(*
SPDX-FileCopyrightText: © 2026 Oleksandr Tiutyk <trofimich@gmail.com>
SPDX-License-Identifier: MIT
License: https://opensource.org/license/mit
*)

(*!
<summary>Creates generic value descriptors by borrowing, adopting or cloning data.</summary>
<description>
Object cloning requires ICloneable; other cloned values are copied as bytes. Owning modes require permission
to release the stored allocation. Exception objects and their engine-managed clones are unsupported in
user-managed generic collections.
</description>
*)

{attribute 'no_explicit_call' := 'do not call this function block directly'}
PROGRAM GenericValueFactory
VAR_OUTPUT
	GenericValueClassName : STRING := 'GENERIC_VALUE';
END_VAR
VAR
	{attribute 'hide'} 
	_ClassName : STRING := __POUNAME();
END_VAR

{attribute 'monitoring' := 'call'}
PROPERTY ClassName : REFERENCE TO STRING
GET
ClassName REF= _ClassName;
END_GET
END_PROPERTY

(*!
<summary>Creates a generic descriptor from runtime type metadata and the requested memory policy.</summary>
<description>
TYPE_ENUM and TYPE_SUBRANGE are interpreted as unsigned integers of the same byte size; their signedness and
original type identity are not retained. Convert explicitly to a signed integer first when signed numeric
meaning is required. Borrowing a converted variable references that variable, not the original enum/subrange.
The selected memory policy and cloning requirements follow FromParts; borrowed storage must remain alive while
used.
</description>
*)
METHOD FromAny : GENERIC_VALUE
VAR_INPUT
	value : ANY;
	isObject : BOOL;
	memoryManagementBehavior : GENERIC_MEMORY_MANAGEMENT_BEHAVIOR;
END_VAR
FromAny := FromAnyType(
	value := value,
	isObject := isObject,
	memoryManagementBehavior := memoryManagementBehavior
);
END_METHOD

(*!
<summary>Creates a generic descriptor from runtime type metadata and the requested memory policy.</summary>
<description>
TYPE_ENUM and TYPE_SUBRANGE are interpreted as unsigned integers of the same byte size; their signedness and
original type identity are not retained. Convert explicitly to a signed integer first when signed numeric
meaning is required. Borrowing a converted variable references that variable, not the original enum/subrange.
The selected memory policy and cloning requirements follow FromParts; borrowed storage must remain alive while
used.
</description>
*)
METHOD FromAnyType : GENERIC_VALUE
VAR_INPUT
	value : __SYSTEM.AnyType;
	isObject : BOOL;
	memoryManagementBehavior : GENERIC_MEMORY_MANAGEMENT_BEHAVIOR;
END_VAR
FromAnyType := FromParts(
        	genericTypeClass := GenericTypeClassConvertor.GetGenericTypeClassBySystemAnyType(systemAnyType := value, isObject := isObject),
        	address := value.pValue,
        	size := TO_ULINT(value.diSize),
        	memoryManagementBehavior := memoryManagementBehavior
        );
END_METHOD

(*!
<summary>Borrows existing storage as a BOOLEAN descriptor.</summary>
<description>
Does not copy or own the payload. The caller keeps the source alive and its representation stable while the
descriptor is used. Size is the byte size of the source variable.
</description>
*)
METHOD FromBoolReference : GENERIC_VALUE
VAR_IN_OUT
	value : BOOL;
END_VAR
FromBoolReference := FromParts(
        	genericTypeClass := GENERIC_TYPE_CLASS.BOOLEAN,
        	address := ADR(value),
        	size := XSIZEOF(value),
        	memoryManagementBehavior := GENERIC_MEMORY_MANAGEMENT_BEHAVIOR.STORE_ORIGINAL_REFERENCE_AND_NOT_OWNS_MEMORY
        );
END_METHOD

(*!
<summary>Creates an owned snapshot of a BOOL value.</summary>
<description>
The result is independent of the input storage; release it or transfer ownership exactly once. Allocation
failure uses the framework terminal allocation path. Uses FromAny cloning; the source value is not modified.
</description>
*)
METHOD FromBoolValue : GENERIC_VALUE
VAR_INPUT
	value : BOOL;
END_VAR
FromBoolValue := FromAny(
	value := value,
	isObject := FALSE,
	memoryManagementBehavior := GENERIC_MEMORY_MANAGEMENT_BEHAVIOR.CLONE_ORIGINAL_VALUE_AND_OWNS_MEMORY
);
END_METHOD

(*!
<summary>Borrows existing storage as a UINT_8 descriptor.</summary>
<description>
Does not copy or own the payload. The caller keeps the source alive and its representation stable while the
descriptor is used. Size is the byte size of the source variable.
</description>
*)
METHOD FromByteReference : GENERIC_VALUE
VAR_IN_OUT
	value : BYTE;
END_VAR
FromByteReference := FromParts(
        	genericTypeClass := GENERIC_TYPE_CLASS.UINT_8,
        	address := ADR(value),
        	size := XSIZEOF(value),
        	memoryManagementBehavior := GENERIC_MEMORY_MANAGEMENT_BEHAVIOR.STORE_ORIGINAL_REFERENCE_AND_NOT_OWNS_MEMORY
        );
END_METHOD

(*!
<summary>Creates an owned snapshot of a BYTE value.</summary>
<description>
The result is independent of the input storage; release it or transfer ownership exactly once. Allocation
failure uses the framework terminal allocation path. Uses FromAny cloning; the source value is not modified.
</description>
*)
METHOD FromByteValue : GENERIC_VALUE
VAR_INPUT
	value : BYTE;
END_VAR
FromByteValue := FromAny(
	value := value,
	isObject := FALSE,
	memoryManagementBehavior := GENERIC_MEMORY_MANAGEMENT_BEHAVIOR.CLONE_ORIGINAL_VALUE_AND_OWNS_MEMORY
);
END_METHOD

(*!
<summary>Borrows existing storage as a DATE_AND_TIME_32 descriptor.</summary>
<description>
Does not copy or own the payload. The caller keeps the source alive and its representation stable while the
descriptor is used. Size is the byte size of the source variable.
</description>
*)
METHOD FromDateAndTimeReference : GENERIC_VALUE
VAR_IN_OUT
	value : DATE_AND_TIME;
END_VAR
FromDateAndTimeReference := FromParts(
        	genericTypeClass := GENERIC_TYPE_CLASS.DATE_AND_TIME_32,
        	address := ADR(value),
        	size := XSIZEOF(value),
        	memoryManagementBehavior := GENERIC_MEMORY_MANAGEMENT_BEHAVIOR.STORE_ORIGINAL_REFERENCE_AND_NOT_OWNS_MEMORY
        );
END_METHOD

(*!
<summary>Creates an owned snapshot of a DATE_AND_TIME value.</summary>
<description>
The result is independent of the input storage; release it or transfer ownership exactly once. Allocation
failure uses the framework terminal allocation path. Uses FromAny cloning; the source value is not modified.
</description>
*)
METHOD FromDateAndTimeValue : GENERIC_VALUE
VAR_INPUT
	value : DATE_AND_TIME;
END_VAR
FromDateAndTimeValue := FromAny(
	value := value,
	isObject := FALSE,
	memoryManagementBehavior := GENERIC_MEMORY_MANAGEMENT_BEHAVIOR.CLONE_ORIGINAL_VALUE_AND_OWNS_MEMORY
);
END_METHOD

(*!
<summary>Borrows existing storage as a DATE_32 descriptor.</summary>
<description>
Does not copy or own the payload. The caller keeps the source alive and its representation stable while the
descriptor is used. Size is the byte size of the source variable.
</description>
*)
METHOD FromDateReference : GENERIC_VALUE
VAR_IN_OUT
	value : DATE;
END_VAR
FromDateReference := FromParts(
        	genericTypeClass := GENERIC_TYPE_CLASS.DATE_32,
        	address := ADR(value),
        	size := XSIZEOF(value),
        	memoryManagementBehavior := GENERIC_MEMORY_MANAGEMENT_BEHAVIOR.STORE_ORIGINAL_REFERENCE_AND_NOT_OWNS_MEMORY
        );
END_METHOD

(*!
<summary>Creates an owned snapshot of a DATE value.</summary>
<description>
The result is independent of the input storage; release it or transfer ownership exactly once. Allocation
failure uses the framework terminal allocation path. Uses FromAny cloning; the source value is not modified.
</description>
*)
METHOD FromDateValue : GENERIC_VALUE
VAR_INPUT
	value : DATE;
END_VAR
FromDateValue := FromAny(
	value := value,
	isObject := FALSE,
	memoryManagementBehavior := GENERIC_MEMORY_MANAGEMENT_BEHAVIOR.CLONE_ORIGINAL_VALUE_AND_OWNS_MEMORY
);
END_METHOD

(*!
<summary>Borrows existing storage as a INT_32 descriptor.</summary>
<description>
Does not copy or own the payload. The caller keeps the source alive and its representation stable while the
descriptor is used. Size is the byte size of the source variable.
</description>
*)
METHOD FromDIntReference : GENERIC_VALUE
VAR_IN_OUT
	value : DINT;
END_VAR
FromDIntReference := FromParts(
        	genericTypeClass := GENERIC_TYPE_CLASS.INT_32,
        	address := ADR(value),
        	size := XSIZEOF(value),
        	memoryManagementBehavior := GENERIC_MEMORY_MANAGEMENT_BEHAVIOR.STORE_ORIGINAL_REFERENCE_AND_NOT_OWNS_MEMORY
        );
END_METHOD

(*!
<summary>Creates an owned snapshot of a DINT value.</summary>
<description>
The result is independent of the input storage; release it or transfer ownership exactly once. Allocation
failure uses the framework terminal allocation path. Uses FromAny cloning; the source value is not modified.
</description>
*)
METHOD FromDIntValue : GENERIC_VALUE
VAR_INPUT
	value : DINT;
END_VAR
FromDIntValue := FromAny(
	value := value,
	isObject := FALSE,
	memoryManagementBehavior := GENERIC_MEMORY_MANAGEMENT_BEHAVIOR.CLONE_ORIGINAL_VALUE_AND_OWNS_MEMORY
);
END_METHOD

(*!
<summary>Borrows existing storage as a UINT_32 descriptor.</summary>
<description>
Does not copy or own the payload. The caller keeps the source alive and its representation stable while the
descriptor is used. Size is the byte size of the source variable.
</description>
*)
METHOD FromDWordReference : GENERIC_VALUE
VAR_IN_OUT
	value : DWORD;
END_VAR
FromDWordReference := FromParts(
        	genericTypeClass := GENERIC_TYPE_CLASS.UINT_32,
        	address := ADR(value),
        	size := XSIZEOF(value),
        	memoryManagementBehavior := GENERIC_MEMORY_MANAGEMENT_BEHAVIOR.STORE_ORIGINAL_REFERENCE_AND_NOT_OWNS_MEMORY
        );
END_METHOD

(*!
<summary>Creates an owned snapshot of a DWORD value.</summary>
<description>
The result is independent of the input storage; release it or transfer ownership exactly once. Allocation
failure uses the framework terminal allocation path. Uses FromAny cloning; the source value is not modified.
</description>
*)
METHOD FromDWordValue : GENERIC_VALUE
VAR_INPUT
	value : DWORD;
END_VAR
FromDWordValue := FromAny(
	value := value,
	isObject := FALSE,
	memoryManagementBehavior := GENERIC_MEMORY_MANAGEMENT_BEHAVIOR.CLONE_ORIGINAL_VALUE_AND_OWNS_MEMORY
);
END_METHOD

(*!
<summary>Borrows existing storage as a INT_16 descriptor.</summary>
<description>
Does not copy or own the payload. The caller keeps the source alive and its representation stable while the
descriptor is used. Size is the byte size of the source variable.
</description>
*)
METHOD FromIntReference : GENERIC_VALUE
VAR_IN_OUT
	value : INT;
END_VAR
FromIntReference := FromParts(
        	genericTypeClass := GENERIC_TYPE_CLASS.INT_16,
        	address := ADR(value),
        	size := XSIZEOF(value),
        	memoryManagementBehavior := GENERIC_MEMORY_MANAGEMENT_BEHAVIOR.STORE_ORIGINAL_REFERENCE_AND_NOT_OWNS_MEMORY
        );
END_METHOD

(*!
<summary>Creates an owned snapshot of a INT value.</summary>
<description>
The result is independent of the input storage; release it or transfer ownership exactly once. Allocation
failure uses the framework terminal allocation path. Uses FromAny cloning; the source value is not modified.
</description>
*)
METHOD FromIntValue : GENERIC_VALUE
VAR_INPUT
	value : INT;
END_VAR
FromIntValue := FromAny(
	value := value,
	isObject := FALSE,
	memoryManagementBehavior := GENERIC_MEMORY_MANAGEMENT_BEHAVIOR.CLONE_ORIGINAL_VALUE_AND_OWNS_MEMORY
);
END_METHOD

(*!
<summary>Creates a non-owning descriptor for an existing object.</summary>
<description>
Null input raises ArgumentNotSpecifiedException. Uses the live object SelfAddress and SelfSize; does not clone
or retain ownership. The object must outlive all uses of the result.
</description>
*)
METHOD FromIObjectReference : GENERIC_VALUE
VAR_INPUT
	instance : IObject;
END_VAR
IF instance = 0 THEN
	Exceptions.ThrowArgumentNotSpecified(
		sourceNamespaceName := NamespaceName,
		sourceClassName := ClassName,
		sourcePOUName := __POUNAME(),
		sourcePosition := __POSITION(),
		argumentName := 'instance'
	);
END_IF

FromIObjectReference := FromParts(
		genericTypeClass := GENERIC_TYPE_CLASS.OBJECT,
		address := instance.SelfAddress,
		size := instance.SelfSize,
		memoryManagementBehavior := GENERIC_MEMORY_MANAGEMENT_BEHAVIOR.STORE_ORIGINAL_REFERENCE_AND_NOT_OWNS_MEMORY
	);
END_METHOD

(*!
<summary>Creates an owning descriptor for a clone of an object.</summary>
<description>
Null input raises ArgumentNotSpecifiedException. Uses the FromParts object-clone contract: a suitable
independent ICloneable result is required; failure raises an exception. The caller must release or transfer
the result exactly once. Task-managed exception clones are not supported as owned generic values.
</description>
*)
METHOD FromIObjectValue : GENERIC_VALUE 
VAR_INPUT
	instance : IObject;
END_VAR
IF instance = 0 THEN
	Exceptions.ThrowArgumentNotSpecified(
		sourceNamespaceName := NamespaceName,
		sourceClassName := ClassName,
		sourcePOUName := __POUNAME(),
		sourcePosition := __POSITION(),
		argumentName := 'instance'
	);
END_IF

FromIObjectValue := FromParts(
		genericTypeClass := GENERIC_TYPE_CLASS.OBJECT,
		address := instance.SelfAddress,
		size := instance.SelfSize,
		memoryManagementBehavior := GENERIC_MEMORY_MANAGEMENT_BEHAVIOR.CLONE_ORIGINAL_VALUE_AND_OWNS_MEMORY
	);
END_METHOD

(*!
<summary>Creates a borrowed generic descriptor for an LDATE_AND_TIME variable.</summary>
<description>
Preserves the DATE_AND_TIME_64 category and references the original variable without copying or allocating
storage. The caller keeps the variable alive while the descriptor is used; ownership is not transferred.
</description>
*)
//!<param name="value">Variable whose storage is borrowed by the returned descriptor.</param>
METHOD FromLDateAndTimeReference : GENERIC_VALUE
VAR_IN_OUT
	value : LDATE_AND_TIME;
END_VAR
FromLDateAndTimeReference := FromParts(
        	genericTypeClass := GENERIC_TYPE_CLASS.DATE_AND_TIME_64,
        	address := ADR(value),
        	size := XSIZEOF(value),
        	memoryManagementBehavior := GENERIC_MEMORY_MANAGEMENT_BEHAVIOR.STORE_ORIGINAL_REFERENCE_AND_NOT_OWNS_MEMORY
        );
END_METHOD

(*!
<summary>Creates an owned snapshot of a LDATE_AND_TIME value.</summary>
<description>
The result is independent of the input storage; release it or transfer ownership exactly once. Allocation
failure uses the framework terminal allocation path. Uses FromAny cloning; the source value is not modified.
</description>
*)
METHOD FromLDateAndTimeValue : GENERIC_VALUE
VAR_INPUT
	value : LDATE_AND_TIME;
END_VAR
FromLDateAndTimeValue := FromAny(
	value := value,
	isObject := FALSE,
	memoryManagementBehavior := GENERIC_MEMORY_MANAGEMENT_BEHAVIOR.CLONE_ORIGINAL_VALUE_AND_OWNS_MEMORY
);
END_METHOD

(*!
<summary>Creates a borrowed generic descriptor for an LDATE variable.</summary>
<description>
Preserves the DATE_64 category and references the original variable without copying or allocating storage. The
caller keeps the variable alive while the descriptor is used; ownership is not transferred.
</description>
*)
//!<param name="value">Variable whose storage is borrowed by the returned descriptor.</param>
METHOD FromLDateReference : GENERIC_VALUE
VAR_IN_OUT
	value : LDATE;
END_VAR
FromLDateReference := FromParts(
        	genericTypeClass := GENERIC_TYPE_CLASS.DATE_64,
        	address := ADR(value),
        	size := XSIZEOF(value),
        	memoryManagementBehavior := GENERIC_MEMORY_MANAGEMENT_BEHAVIOR.STORE_ORIGINAL_REFERENCE_AND_NOT_OWNS_MEMORY
        );
END_METHOD

(*!
<summary>Creates an owned snapshot of a LDATE value.</summary>
<description>
The result is independent of the input storage; release it or transfer ownership exactly once. Allocation
failure uses the framework terminal allocation path. Uses FromAny cloning; the source value is not modified.
</description>
*)
METHOD FromLDateValue : GENERIC_VALUE
VAR_INPUT
	value : LDATE;
END_VAR
FromLDateValue := FromAny(
	value := value,
	isObject := FALSE,
	memoryManagementBehavior := GENERIC_MEMORY_MANAGEMENT_BEHAVIOR.CLONE_ORIGINAL_VALUE_AND_OWNS_MEMORY
);
END_METHOD

(*!
<summary>Borrows existing storage as a INT_64 descriptor.</summary>
<description>
Does not copy or own the payload. The caller keeps the source alive and its representation stable while the
descriptor is used. Size is the byte size of the source variable.
</description>
*)
METHOD FromLIntReference : GENERIC_VALUE
VAR_IN_OUT
	value : LINT;
END_VAR
FromLIntReference := FromParts(
        	genericTypeClass := GENERIC_TYPE_CLASS.INT_64,
        	address := ADR(value),
        	size := XSIZEOF(value),
        	memoryManagementBehavior := GENERIC_MEMORY_MANAGEMENT_BEHAVIOR.STORE_ORIGINAL_REFERENCE_AND_NOT_OWNS_MEMORY
        );
END_METHOD

(*!
<summary>Creates an owned snapshot of a LINT value.</summary>
<description>
The result is independent of the input storage; release it or transfer ownership exactly once. Allocation
failure uses the framework terminal allocation path. Uses FromAny cloning; the source value is not modified.
</description>
*)
METHOD FromLIntValue : GENERIC_VALUE
VAR_INPUT
	value : LINT;
END_VAR
FromLIntValue := FromAny(
	value := value,
	isObject := FALSE,
	memoryManagementBehavior := GENERIC_MEMORY_MANAGEMENT_BEHAVIOR.CLONE_ORIGINAL_VALUE_AND_OWNS_MEMORY
);
END_METHOD

(*!
<summary>Borrows existing storage as a REAL_64 descriptor.</summary>
<description>
Does not copy or own the payload. The caller keeps the source alive and its representation stable while the
descriptor is used. Size is the byte size of the source variable.
</description>
*)
METHOD FromLRealReference : GENERIC_VALUE
VAR_IN_OUT
	value : LREAL;
END_VAR
FromLRealReference := FromParts(
        	genericTypeClass := GENERIC_TYPE_CLASS.REAL_64,
        	address := ADR(value),
        	size := XSIZEOF(value),
        	memoryManagementBehavior := GENERIC_MEMORY_MANAGEMENT_BEHAVIOR.STORE_ORIGINAL_REFERENCE_AND_NOT_OWNS_MEMORY
        );
END_METHOD

(*!
<summary>Creates an owned snapshot of a LREAL value.</summary>
<description>
The result is independent of the input storage; release it or transfer ownership exactly once. Allocation
failure uses the framework terminal allocation path. Uses FromAny cloning; the source value is not modified.
</description>
*)
METHOD FromLRealValue : GENERIC_VALUE
VAR_INPUT
	value : LREAL;
END_VAR
FromLRealValue := FromAny(
	value := value,
	isObject := FALSE,
	memoryManagementBehavior := GENERIC_MEMORY_MANAGEMENT_BEHAVIOR.CLONE_ORIGINAL_VALUE_AND_OWNS_MEMORY
);
END_METHOD

(*!
<summary>Creates a borrowed generic descriptor for an LTIME_OF_DAY variable.</summary>
<description>
Preserves the TIME_OF_DAY_64 category and references the original variable without copying or allocating
storage. The caller keeps the variable alive while the descriptor is used; ownership is not transferred.
</description>
*)
//!<param name="value">Variable whose storage is borrowed by the returned descriptor.</param>
METHOD FromLTimeOfDayReference : GENERIC_VALUE
VAR_IN_OUT
	value : LTIME_OF_DAY;
END_VAR
FromLTimeOfDayReference := FromParts(
        	genericTypeClass := GENERIC_TYPE_CLASS.TIME_OF_DAY_64,
        	address := ADR(value),
        	size := XSIZEOF(value),
        	memoryManagementBehavior := GENERIC_MEMORY_MANAGEMENT_BEHAVIOR.STORE_ORIGINAL_REFERENCE_AND_NOT_OWNS_MEMORY
        );
END_METHOD

(*!
<summary>Creates an owned snapshot of a LTIME_OF_DAY value.</summary>
<description>
The result is independent of the input storage; release it or transfer ownership exactly once. Allocation
failure uses the framework terminal allocation path. Uses FromAny cloning; the source value is not modified.
</description>
*)
METHOD FromLTimeOfDayValue : GENERIC_VALUE
VAR_INPUT
	value : LTIME_OF_DAY;
END_VAR
FromLTimeOfDayValue := FromAny(
	value := value,
	isObject := FALSE,
	memoryManagementBehavior := GENERIC_MEMORY_MANAGEMENT_BEHAVIOR.CLONE_ORIGINAL_VALUE_AND_OWNS_MEMORY
);
END_METHOD

(*!
<summary>Creates a borrowed generic descriptor for an LTIME variable.</summary>
<description>
Preserves the TIME_64 category and references the original variable without copying or allocating storage. The
caller keeps the variable alive while the descriptor is used; ownership is not transferred.
</description>
*)
//!<param name="value">Variable whose storage is borrowed by the returned descriptor.</param>
METHOD FromLTimeReference : GENERIC_VALUE
VAR_IN_OUT
	value : LTIME;
END_VAR
FromLTimeReference := FromParts(
        	genericTypeClass := GENERIC_TYPE_CLASS.TIME_64,
        	address := ADR(value),
        	size := XSIZEOF(value),
        	memoryManagementBehavior := GENERIC_MEMORY_MANAGEMENT_BEHAVIOR.STORE_ORIGINAL_REFERENCE_AND_NOT_OWNS_MEMORY
        );
END_METHOD

(*!
<summary>Creates an owned snapshot of a LTIME value.</summary>
<description>
The result is independent of the input storage; release it or transfer ownership exactly once. Allocation
failure uses the framework terminal allocation path. Uses FromAny cloning; the source value is not modified.
</description>
*)
METHOD FromLTimeValue : GENERIC_VALUE
VAR_INPUT
	value : LTIME;
END_VAR
FromLTimeValue := FromAny(
	value := value,
	isObject := FALSE,
	memoryManagementBehavior := GENERIC_MEMORY_MANAGEMENT_BEHAVIOR.CLONE_ORIGINAL_VALUE_AND_OWNS_MEMORY
);
END_METHOD

(*!
<summary>Borrows existing storage as a UINT_64 descriptor.</summary>
<description>
Does not copy or own the payload. The caller keeps the source alive and its representation stable while the
descriptor is used. Size is the byte size of the source variable.
</description>
*)
METHOD FromLWordReference : GENERIC_VALUE
VAR_IN_OUT
	value : LWORD;
END_VAR
FromLWordReference := FromParts(
        	genericTypeClass := GENERIC_TYPE_CLASS.UINT_64,
        	address := ADR(value),
        	size := XSIZEOF(value),
        	memoryManagementBehavior := GENERIC_MEMORY_MANAGEMENT_BEHAVIOR.STORE_ORIGINAL_REFERENCE_AND_NOT_OWNS_MEMORY
        );
END_METHOD

(*!
<summary>Creates an owned snapshot of a LWORD value.</summary>
<description>
The result is independent of the input storage; release it or transfer ownership exactly once. Allocation
failure uses the framework terminal allocation path. Uses FromAny cloning; the source value is not modified.
</description>
*)
METHOD FromLWordValue : GENERIC_VALUE
VAR_INPUT
	value : LWORD;
END_VAR
FromLWordValue := FromAny(
	value := value,
	isObject := FALSE,
	memoryManagementBehavior := GENERIC_MEMORY_MANAGEMENT_BEHAVIOR.CLONE_ORIGINAL_VALUE_AND_OWNS_MEMORY
);
END_METHOD

(*!
<summary>Creates a non-owning descriptor for an existing object.</summary>
<description>
Null input raises ArgumentNotSpecifiedException. Uses the live object SelfAddress and SelfSize; does not clone
or retain ownership. The object must outlive all uses of the result.
</description>
*)
METHOD FromObjectReference : GENERIC_VALUE
VAR_INPUT
	instance : REFERENCE TO Object;
END_VAR
IF NOT __ISVALIDREF(instance) THEN
	Exceptions.ThrowArgumentNotSpecified(
		sourceNamespaceName := NamespaceName,
		sourceClassName := ClassName,
		sourcePOUName := __POUNAME(),
		sourcePosition := __POSITION(),
		argumentName := 'instance'
	);
END_IF

FromObjectReference := FromParts(
		genericTypeClass := GENERIC_TYPE_CLASS.OBJECT,
		address := instance.SelfAddress,
		size := instance.SelfSize,
		memoryManagementBehavior := GENERIC_MEMORY_MANAGEMENT_BEHAVIOR.STORE_ORIGINAL_REFERENCE_AND_NOT_OWNS_MEMORY
	);
END_METHOD

(*!
<summary>Creates an owning generic descriptor for a clone of the supplied object.</summary>
<description>
Requires a live object implementing ICloneable whose clone may be released by the owner of the returned
descriptor. Throws ArgumentNotSpecifiedException for a null reference or NotSupportedException when ICloneable
is absent. The original object is not adopted.
</description>
*)
//!<param name="instance">Object to clone through ICloneable.</param>
METHOD FromObjectValue : GENERIC_VALUE 
VAR_INPUT
	instance : REFERENCE TO Object;
END_VAR
IF NOT __ISVALIDREF(instance) THEN
	Exceptions.ThrowArgumentNotSpecified(
		sourceNamespaceName := NamespaceName,
		sourceClassName := ClassName,
		sourcePOUName := __POUNAME(),
		sourcePosition := __POSITION(),
		argumentName := 'instance'
	);
END_IF

FromObjectValue := FromParts(
		genericTypeClass := GENERIC_TYPE_CLASS.OBJECT,
		address := instance.SelfAddress,
		size := instance.SelfSize,
		memoryManagementBehavior := GENERIC_MEMORY_MANAGEMENT_BEHAVIOR.CLONE_ORIGINAL_VALUE_AND_OWNS_MEMORY
	);
END_METHOD

(*!
<summary>Creates a generic value from a type, address, size and memory-management policy.</summary>
<description>
Owning modes require permission to release the stored allocation, including any result returned by Clone. In
clone mode, OBJECT requires ICloneable; otherwise NotSupportedException is raised. Clone must return a
non-null object on success and raise an exception on failure; its exceptions propagate. Failure to allocate a
byte copy invokes the terminal DynamicMemoryManager.RaiseAllocationFailure mechanism. Other type categories
are copied as bytes, without recursively cloning referenced resources. For a nonempty byte copy, size above
UnsignedInt32.MAX_VALUE raises ArgumentOutOfRangeException before allocation or conversion to UDINT. Exception
objects and their engine-managed clones are not supported by user-managed generic collections. Their lifetime
ends at cycle cleanup; use ERROR to retain an error as state.
</description>
*)
METHOD FromParts : GENERIC_VALUE
VAR_INPUT
	genericTypeClass : GENERIC_TYPE_CLASS;
	address : POINTER TO BYTE;
	size : ULINT;
	memoryManagementBehavior : GENERIC_MEMORY_MANAGEMENT_BEHAVIOR;
END_VAR
VAR
	newAddress : POINTER TO BYTE;

	objectPointer : POINTER TO Object;
	cloneable : ICloneable;
	clone : IObject;

END_VAR
IF address = 0 OR_ELSE size <= 0 THEN
	RETURN;
END_IF

CASE memoryManagementBehavior OF
	GENERIC_MEMORY_MANAGEMENT_BEHAVIOR.CLONE_ORIGINAL_VALUE_AND_OWNS_MEMORY:
		IF genericTypeClass = GENERIC_TYPE_CLASS.OBJECT THEN
			objectPointer := address;

			IF NOT __QUERYINTERFACE(objectPointer^, cloneable) THEN
				Exceptions.ThrowNotSupported(
					sourceNamespaceName := NamespaceName,
					sourceClassName := ClassName,
					sourcePOUName := __POUNAME(),
					sourcePosition := __POSITION(),
					message := "Object cloning requires ICloneable."
				);
			END_IF

			clone := cloneable.Clone();
			newAddress := clone.SelfAddress;	
		ELSE
			IF size > TO_ULINT(UnsignedInt32.MAX_VALUE) THEN
				Exceptions.ThrowArgumentOutOfRange(
					sourceNamespaceName := NamespaceName,
					sourceClassName := ClassName,
					sourcePOUName := __POUNAME(),
					sourcePosition := __POSITION(),
					argumentName := 'size',
					argumentValue := size
				);
			END_IF

			newAddress := __NEW(BYTE, TO_UDINT(size));

			IF newAddress = 0 THEN
				DynamicMemoryManager.RaiseAllocationFailure();
			END_IF

			Tc2_System.MEMCPY(destAddr := newAddress, srcAddr := address, n := TO_UDINT(size));
		END_IF

		FromParts.Assign(genericTypeClass := genericTypeClass, address := newAddress, size := size, isMemoryOwner := TRUE);
	
	GENERIC_MEMORY_MANAGEMENT_BEHAVIOR.STORE_ORIGINAL_REFERENCE_AND_NOT_OWNS_MEMORY:
		FromParts.Assign(genericTypeClass := genericTypeClass, address := address, size := size, isMemoryOwner := FALSE);
	
	GENERIC_MEMORY_MANAGEMENT_BEHAVIOR.STORE_ORIGINAL_REFERENCE_AND_OWNS_MEMORY:
		FromParts.Assign(genericTypeClass := genericTypeClass, address := address, size := size, isMemoryOwner := TRUE);
END_CASE
END_METHOD

(*!
<summary>Borrows existing storage as a REAL_32 descriptor.</summary>
<description>
Does not copy or own the payload. The caller keeps the source alive and its representation stable while the
descriptor is used. Size is the byte size of the source variable.
</description>
*)
METHOD FromRealReference : GENERIC_VALUE
VAR_IN_OUT
	value : REAL;
END_VAR
FromRealReference := FromParts(
        	genericTypeClass := GENERIC_TYPE_CLASS.REAL_32,
        	address := ADR(value),
        	size := XSIZEOF(value),
        	memoryManagementBehavior := GENERIC_MEMORY_MANAGEMENT_BEHAVIOR.STORE_ORIGINAL_REFERENCE_AND_NOT_OWNS_MEMORY
        );
END_METHOD

(*!
<summary>Creates an owned snapshot of a REAL value.</summary>
<description>
The result is independent of the input storage; release it or transfer ownership exactly once. Allocation
failure uses the framework terminal allocation path. Uses FromAny cloning; the source value is not modified.
</description>
*)
METHOD FromRealValue : GENERIC_VALUE
VAR_INPUT
	value : REAL;
END_VAR
FromRealValue := FromAny(
	value := value,
	isObject := FALSE,
	memoryManagementBehavior := GENERIC_MEMORY_MANAGEMENT_BEHAVIOR.CLONE_ORIGINAL_VALUE_AND_OWNS_MEMORY
);
END_METHOD

(*!
<summary>Borrows existing storage as a INT_8 descriptor.</summary>
<description>
Does not copy or own the payload. The caller keeps the source alive and its representation stable while the
descriptor is used. Size is the byte size of the source variable.
</description>
*)
METHOD FromSIntReference : GENERIC_VALUE
VAR_IN_OUT
	value : SINT;
END_VAR
FromSIntReference := FromParts(
        	genericTypeClass := GENERIC_TYPE_CLASS.INT_8,
        	address := ADR(value),
        	size := XSIZEOF(value),
        	memoryManagementBehavior := GENERIC_MEMORY_MANAGEMENT_BEHAVIOR.STORE_ORIGINAL_REFERENCE_AND_NOT_OWNS_MEMORY
        );
END_METHOD

(*!
<summary>Creates an owned snapshot of a SINT value.</summary>
<description>
The result is independent of the input storage; release it or transfer ownership exactly once. Allocation
failure uses the framework terminal allocation path. Uses FromAny cloning; the source value is not modified.
</description>
*)
METHOD FromSIntValue : GENERIC_VALUE
VAR_INPUT
	value : SINT;
END_VAR
FromSIntValue := FromAny(
	value := value,
	isObject := FALSE,
	memoryManagementBehavior := GENERIC_MEMORY_MANAGEMENT_BEHAVIOR.CLONE_ORIGINAL_VALUE_AND_OWNS_MEMORY
);
END_METHOD

(*!
<summary>Borrows existing storage as a STRING_8 descriptor.</summary>
<description>
Does not copy or own the payload. The caller keeps the source alive and its representation stable while the
descriptor is used. Size records the current text including its terminator, not the full declared buffer
capacity.
</description>
*)
METHOD FromStringReference : GENERIC_VALUE
VAR_IN_OUT CONSTANT
	value : STRING;
END_VAR
FromStringReference := FromParts(
	genericTypeClass := GENERIC_TYPE_CLASS.STRING_8,
	address := ADR(value),
	size := Strings.GetActualSize(value := value),
	memoryManagementBehavior := GENERIC_MEMORY_MANAGEMENT_BEHAVIOR.STORE_ORIGINAL_REFERENCE_AND_NOT_OWNS_MEMORY
);
END_METHOD

(*!
<summary>Creates an owned snapshot of a STRING value.</summary>
<description>
The result is independent of the input storage; release it or transfer ownership exactly once. Allocation
failure uses the framework terminal allocation path. Copies current text including its terminator, not unused
buffer capacity.
</description>
*)
METHOD FromStringValue : GENERIC_VALUE
VAR_IN_OUT CONSTANT
	value : STRING;
END_VAR
FromStringValue := FromParts(
        	genericTypeClass := GENERIC_TYPE_CLASS.STRING_8,
        	address := ADR(value),
        	size := Strings.GetActualSize(value := value),
        	memoryManagementBehavior := GENERIC_MEMORY_MANAGEMENT_BEHAVIOR.CLONE_ORIGINAL_VALUE_AND_OWNS_MEMORY
        );
END_METHOD

(*!
<summary>Borrows existing storage as a TIME_OF_DAY_32 descriptor.</summary>
<description>
Does not copy or own the payload. The caller keeps the source alive and its representation stable while the
descriptor is used. Size is the byte size of the source variable.
</description>
*)
METHOD FromTimeOfDayReference : GENERIC_VALUE
VAR_IN_OUT
	value : TIME_OF_DAY;
END_VAR
FromTimeOfDayReference := FromParts(
        	genericTypeClass := GENERIC_TYPE_CLASS.TIME_OF_DAY_32,
        	address := ADR(value),
        	size := XSIZEOF(value),
        	memoryManagementBehavior := GENERIC_MEMORY_MANAGEMENT_BEHAVIOR.STORE_ORIGINAL_REFERENCE_AND_NOT_OWNS_MEMORY
        );
END_METHOD

(*!
<summary>Creates an owned snapshot of a TIME_OF_DAY value.</summary>
<description>
The result is independent of the input storage; release it or transfer ownership exactly once. Allocation
failure uses the framework terminal allocation path. Uses FromAny cloning; the source value is not modified.
</description>
*)
METHOD FromTimeOfDayValue : GENERIC_VALUE
VAR_INPUT
	value : TIME_OF_DAY;
END_VAR
FromTimeOfDayValue := FromAny(
	value := value,
	isObject := FALSE,
	memoryManagementBehavior := GENERIC_MEMORY_MANAGEMENT_BEHAVIOR.CLONE_ORIGINAL_VALUE_AND_OWNS_MEMORY
);
END_METHOD

(*!
<summary>Borrows existing storage as a TIME_32 descriptor.</summary>
<description>
Does not copy or own the payload. The caller keeps the source alive and its representation stable while the
descriptor is used. Size is the byte size of the source variable.
</description>
*)
METHOD FromTimeReference : GENERIC_VALUE
VAR_IN_OUT
	value : TIME;
END_VAR
FromTimeReference := FromParts(
        	genericTypeClass := GENERIC_TYPE_CLASS.TIME_32,
        	address := ADR(value),
        	size := XSIZEOF(value),
        	memoryManagementBehavior := GENERIC_MEMORY_MANAGEMENT_BEHAVIOR.STORE_ORIGINAL_REFERENCE_AND_NOT_OWNS_MEMORY
        );
END_METHOD

(*!
<summary>Creates an owned snapshot of a TIME value.</summary>
<description>
The result is independent of the input storage; release it or transfer ownership exactly once. Allocation
failure uses the framework terminal allocation path. Uses FromAny cloning; the source value is not modified.
</description>
*)
METHOD FromTimeValue : GENERIC_VALUE
VAR_INPUT
	value : TIME;
END_VAR
FromTimeValue := FromAny(
	value := value,
	isObject := FALSE,
	memoryManagementBehavior := GENERIC_MEMORY_MANAGEMENT_BEHAVIOR.CLONE_ORIGINAL_VALUE_AND_OWNS_MEMORY
);
END_METHOD

(*!
<summary>Borrows existing storage as a UINT_32 descriptor.</summary>
<description>
Does not copy or own the payload. The caller keeps the source alive and its representation stable while the
descriptor is used. Size is the byte size of the source variable.
</description>
*)
METHOD FromUDIntReference : GENERIC_VALUE
VAR_IN_OUT
	value : UDINT;
END_VAR
FromUDIntReference := FromParts(
        	genericTypeClass := GENERIC_TYPE_CLASS.UINT_32,
        	address := ADR(value),
        	size := XSIZEOF(value),
        	memoryManagementBehavior := GENERIC_MEMORY_MANAGEMENT_BEHAVIOR.STORE_ORIGINAL_REFERENCE_AND_NOT_OWNS_MEMORY
        );
END_METHOD

(*!
<summary>Creates an owned snapshot of a UDINT value.</summary>
<description>
The result is independent of the input storage; release it or transfer ownership exactly once. Allocation
failure uses the framework terminal allocation path. Uses FromAny cloning; the source value is not modified.
</description>
*)
METHOD FromUDIntValue : GENERIC_VALUE
VAR_INPUT
	value : UDINT;
END_VAR
FromUDIntValue := FromAny(
	value := value,
	isObject := FALSE,
	memoryManagementBehavior := GENERIC_MEMORY_MANAGEMENT_BEHAVIOR.CLONE_ORIGINAL_VALUE_AND_OWNS_MEMORY
);
END_METHOD

(*!
<summary>Borrows existing storage as a UINT_16 descriptor.</summary>
<description>
Does not copy or own the payload. The caller keeps the source alive and its representation stable while the
descriptor is used. Size is the byte size of the source variable.
</description>
*)
METHOD FromUIntReference : GENERIC_VALUE
VAR_IN_OUT
	value : UINT;
END_VAR
FromUIntReference := FromParts(
        	genericTypeClass := GENERIC_TYPE_CLASS.UINT_16,
        	address := ADR(value),
        	size := XSIZEOF(value),
        	memoryManagementBehavior := GENERIC_MEMORY_MANAGEMENT_BEHAVIOR.STORE_ORIGINAL_REFERENCE_AND_NOT_OWNS_MEMORY
        );
END_METHOD

(*!
<summary>Creates an owned snapshot of a UINT value.</summary>
<description>
The result is independent of the input storage; release it or transfer ownership exactly once. Allocation
failure uses the framework terminal allocation path. Uses FromAny cloning; the source value is not modified.
</description>
*)
METHOD FromUIntValue : GENERIC_VALUE
VAR_INPUT
	value : UINT;
END_VAR
FromUIntValue := FromAny(
	value := value,
	isObject := FALSE,
	memoryManagementBehavior := GENERIC_MEMORY_MANAGEMENT_BEHAVIOR.CLONE_ORIGINAL_VALUE_AND_OWNS_MEMORY
);
END_METHOD

(*!
<summary>Borrows existing storage as a UINT_64 descriptor.</summary>
<description>
Does not copy or own the payload. The caller keeps the source alive and its representation stable while the
descriptor is used. Size is the byte size of the source variable.
</description>
*)
METHOD FromULIntReference : GENERIC_VALUE
VAR_IN_OUT
	value : ULINT;
END_VAR
FromULIntReference := FromParts(
        	genericTypeClass := GENERIC_TYPE_CLASS.UINT_64,
        	address := ADR(value),
        	size := XSIZEOF(value),
        	memoryManagementBehavior := GENERIC_MEMORY_MANAGEMENT_BEHAVIOR.STORE_ORIGINAL_REFERENCE_AND_NOT_OWNS_MEMORY
        );
END_METHOD

(*!
<summary>Creates an owned snapshot of a ULINT value.</summary>
<description>
The result is independent of the input storage; release it or transfer ownership exactly once. Allocation
failure uses the framework terminal allocation path. Uses FromAny cloning; the source value is not modified.
</description>
*)
METHOD FromULIntValue : GENERIC_VALUE
VAR_INPUT
	value : ULINT;
END_VAR
FromULIntValue := FromAny(
	value := value,
	isObject := FALSE,
	memoryManagementBehavior := GENERIC_MEMORY_MANAGEMENT_BEHAVIOR.CLONE_ORIGINAL_VALUE_AND_OWNS_MEMORY
);
END_METHOD

(*!
<summary>Borrows existing storage as a UINT_8 descriptor.</summary>
<description>
Does not copy or own the payload. The caller keeps the source alive and its representation stable while the
descriptor is used. Size is the byte size of the source variable.
</description>
*)
METHOD FromUSIntReference : GENERIC_VALUE
VAR_IN_OUT
	value : USINT;
END_VAR
FromUSIntReference := FromParts(
        	genericTypeClass := GENERIC_TYPE_CLASS.UINT_8,
        	address := ADR(value),
        	size := XSIZEOF(value),
        	memoryManagementBehavior := GENERIC_MEMORY_MANAGEMENT_BEHAVIOR.STORE_ORIGINAL_REFERENCE_AND_NOT_OWNS_MEMORY
        );
END_METHOD

(*!
<summary>Creates an owned snapshot of a USINT value.</summary>
<description>
The result is independent of the input storage; release it or transfer ownership exactly once. Allocation
failure uses the framework terminal allocation path. Uses FromAny cloning; the source value is not modified.
</description>
*)
METHOD FromUSIntValue : GENERIC_VALUE
VAR_INPUT
	value : USINT;
END_VAR
FromUSIntValue := FromAny(
	value := value,
	isObject := FALSE,
	memoryManagementBehavior := GENERIC_MEMORY_MANAGEMENT_BEHAVIOR.CLONE_ORIGINAL_VALUE_AND_OWNS_MEMORY
);
END_METHOD

(*!
<summary>Borrows existing storage as a UINT_16 descriptor.</summary>
<description>
Does not copy or own the payload. The caller keeps the source alive and its representation stable while the
descriptor is used. Size is the byte size of the source variable.
</description>
*)
METHOD FromWordReference : GENERIC_VALUE
VAR_IN_OUT
	value : WORD;
END_VAR
FromWordReference := FromParts(
        	genericTypeClass := GENERIC_TYPE_CLASS.UINT_16,
        	address := ADR(value),
        	size := XSIZEOF(value),
        	memoryManagementBehavior := GENERIC_MEMORY_MANAGEMENT_BEHAVIOR.STORE_ORIGINAL_REFERENCE_AND_NOT_OWNS_MEMORY
        );
END_METHOD

(*!
<summary>Creates an owned snapshot of a WORD value.</summary>
<description>
The result is independent of the input storage; release it or transfer ownership exactly once. Allocation
failure uses the framework terminal allocation path. Uses FromAny cloning; the source value is not modified.
</description>
*)
METHOD FromWordValue : GENERIC_VALUE
VAR_INPUT
	value : WORD;
END_VAR
FromWordValue := FromAny(
	value := value,
	isObject := FALSE,
	memoryManagementBehavior := GENERIC_MEMORY_MANAGEMENT_BEHAVIOR.CLONE_ORIGINAL_VALUE_AND_OWNS_MEMORY
);
END_METHOD

(*!
<summary>Borrows existing storage as a STRING_16 descriptor.</summary>
<description>
Does not copy or own the payload. The caller keeps the source alive and its representation stable while the
descriptor is used. Size records the current text including its terminator, not the full declared buffer
capacity.
</description>
*)
METHOD FromWStringReference : GENERIC_VALUE
VAR_IN_OUT CONSTANT
	value : WSTRING;
END_VAR
FromWStringReference := FromParts(
	genericTypeClass := GENERIC_TYPE_CLASS.STRING_16,
	address := ADR(value),
	size := WideStrings.GetActualSize(value := value),
	memoryManagementBehavior := GENERIC_MEMORY_MANAGEMENT_BEHAVIOR.STORE_ORIGINAL_REFERENCE_AND_NOT_OWNS_MEMORY
);
END_METHOD

(*!
<summary>Creates an owned snapshot of a WSTRING value.</summary>
<description>
The result is independent of the input storage; release it or transfer ownership exactly once. Allocation
failure uses the framework terminal allocation path. Copies current text including its terminator, not unused
buffer capacity.
</description>
*)
METHOD FromWStringValue : GENERIC_VALUE
VAR_IN_OUT CONSTANT
	value : WSTRING;
END_VAR
FromWStringValue := FromParts(
        	genericTypeClass := GENERIC_TYPE_CLASS.STRING_16,
        	address := ADR(value),
        	size := WideStrings.GetActualSize(value := value),
        	memoryManagementBehavior := GENERIC_MEMORY_MANAGEMENT_BEHAVIOR.CLONE_ORIGINAL_VALUE_AND_OWNS_MEMORY
        );
END_METHOD

(*!
<summary>Provides the library namespace used in diagnostics.</summary>
<description>
Borrowed read-only reference to the compiler-initialized library namespace; no ownership transfer.
</description>
*)
{attribute 'monitoring' := 'call'}
PROPERTY NamespaceName : REFERENCE TO STRING
GET
NamespaceName REF= CurrentNamespace.Name;
END_GET
END_PROPERTY

END_PROGRAM

(* stored: Version 1.1.0.1
   POU GenericValueFactory: Id {5aafca66-5cdb-4882-83ad-05bcd6342c33}, SpecialFunc None
   Folder FromTypedReferences: Id {6a62176f-75b8-40f9-88f4-26d2c66b2b4c}
   Folder Date and time: Id {50be7849-3dc1-473b-9a05-6b6e31d6af8b}
   Folder Floating point: Id {135cf303-d7c8-4cb2-83e4-8818dc564814}
   Folder Integer: Id {9822276d-d405-467b-913a-d88d688e27ab}
   Folder Signed: Id {88769d57-d90b-4d86-a952-5ee7177698c2}
   Folder Unsugned: Id {b4e483f8-ba35-4ef4-8231-cc40ee080b19}
   Folder Strings: Id {eee688c5-eebb-4825-a4d2-c0399523c8d1}
   Folder FromTypedValues: Id {25ae72e5-a435-4f95-b7ff-4fa29bd648e4}
   Folder Date and time: Id {c40440d3-8031-4729-9442-ab1c6e1a88ce}
   Folder Floating point: Id {87a9bf3e-1364-4eb7-acac-0cdf6af21cc8}
   Folder Integer: Id {0a1aa935-644b-4556-94c3-416eb3400fa0}
   Folder Signed: Id {940b3a7d-41f9-44cf-8d1e-ff10f12d8a45}
   Folder Unsugned: Id {0879f3ef-e520-4036-bc27-14c1b4a89e4e}
   Folder Strings: Id {b9fa53fd-8c54-4f18-b477-b593285e3922}
   Property ClassName: Id {471a3424-a03f-46e9-aa5d-47ddfd6d5482}
   Get Get: Id {a20ec758-d80c-4890-b9c6-9d76856ede75}
   Method FromAny: Id {6ea8f682-f65a-4f72-b981-df5fc5f1ef43}
   Method FromAnyType: Id {58f5fed2-ee58-4bb7-b5fb-7380db0fc95f}
   Method FromBoolReference: Id {d27b6912-bb8f-448c-b703-74f93763bb2a}
   Method FromBoolValue: Id {05323a56-8230-4256-ab0d-6fb067ae3a7c}
   Method FromByteReference: Id {d0163973-28dc-453e-ad54-13cb227a8692}
   Method FromByteValue: Id {c850b1be-a21b-48c4-b41a-36d350dde20f}
   Method FromDateAndTimeReference: Id {173ac213-1cc9-43cb-af55-055a2d088a5d}
   Method FromDateAndTimeValue: Id {acb7264d-a9f1-46b1-a8df-1b273f60647d}
   Method FromDateReference: Id {e4aa20a7-899e-4891-8b7b-4b75565ece84}
   Method FromDateValue: Id {23c94b95-80f9-479f-a2c5-e7d679fc27d6}
   Method FromDIntReference: Id {347f607f-2c78-4202-8506-027cbef4c70e}
   Method FromDIntValue: Id {3180b989-96c3-434b-b481-bd0a4f94dfea}
   Method FromDWordReference: Id {946efa8e-2ab5-43b1-bf77-3303cffc04cb}
   Method FromDWordValue: Id {a4f9425d-c238-4587-bc3b-6ca752d58eb9}
   Method FromIntReference: Id {297f6b14-cf53-4dfc-8218-a8424a5edfe0}
   Method FromIntValue: Id {8dbf331d-d65d-4447-810a-b5722dd5340b}
   Method FromIObjectReference: Id {5e9ad193-b039-42bb-8395-af4a1c647cfc}
   Method FromIObjectValue: Id {fef270e2-21e0-469c-8151-9d5a311dfd4b}
   Method FromLDateAndTimeReference: Id {73c19958-a0a7-4e2d-ade2-e984449c3d1d}
   Method FromLDateAndTimeValue: Id {a766e905-b94b-4c9d-82d2-dc889e57d0b8}
   Method FromLDateReference: Id {580e428d-fb4b-4375-874d-309e30a280bf}
   Method FromLDateValue: Id {3521f0fd-d786-4c9e-9852-33d078c765f7}
   Method FromLIntReference: Id {3587c5a4-e047-430d-a163-142a19047459}
   Method FromLIntValue: Id {60a27329-0eea-455a-849b-eb1a0f8b3d54}
   Method FromLRealReference: Id {b3eac24c-b062-484b-ad9a-bc37b94b04ce}
   Method FromLRealValue: Id {3dd0d52e-c433-4065-9057-391e0b5d7161}
   Method FromLTimeOfDayReference: Id {ddcd78a1-0fee-4add-a56e-178a6a711394}
   Method FromLTimeOfDayValue: Id {383c7178-c7ae-4a60-9f1e-7d0d454ddfe1}
   Method FromLTimeReference: Id {09bff33e-4edf-4b18-8976-6a561c6f9e70}
   Method FromLTimeValue: Id {720ca242-94c2-488a-8631-0658baa256f2}
   Method FromLWordReference: Id {f772b6da-0878-4a66-aae9-b922e2dd49f9}
   Method FromLWordValue: Id {1b4080c1-48c3-4e24-89fd-b9ed03b1ebe8}
   Method FromObjectReference: Id {1f38a672-fb8f-436c-9ddd-df1d9f011e0c}
   Method FromObjectValue: Id {ad024805-1158-4b96-998d-e6f1c85f0eb0}
   Method FromParts: Id {759e0037-660d-404f-8404-ca0ffa255f71}
   Method FromRealReference: Id {3b55838d-58fe-4935-bf92-dcc94945943e}
   Method FromRealValue: Id {f5d5afa5-da33-48d8-929b-a1880a20b6ed}
   Method FromSIntReference: Id {dcbeabb7-7a7d-43d2-8ece-e53719a456af}
   Method FromSIntValue: Id {69dc6169-e00d-4a1b-a310-c30817210f3f}
   Method FromStringReference: Id {ab2c82b3-b73e-4926-9fa1-21180356ffa0}
   Method FromStringValue: Id {a2ca4991-d75a-4278-817b-66b69acc26fd}
   Method FromTimeOfDayReference: Id {16667815-ae24-4a2e-bb7e-13b02852bf9b}
   Method FromTimeOfDayValue: Id {e882c6af-473d-4d99-a60c-86a44c55080d}
   Method FromTimeReference: Id {4efbab6a-08c6-45a2-8741-5970c5b4615c}
   Method FromTimeValue: Id {9ee9b713-8171-4acb-a940-5ccce35b7698}
   Method FromUDIntReference: Id {1c502058-ad42-4bc4-99e4-7e76741e1405}
   Method FromUDIntValue: Id {168c3430-037e-43ee-96ec-29f9d4ddb82b}
   Method FromUIntReference: Id {81d69bd9-3d0f-4fa9-a701-f3d6b82d40a5}
   Method FromUIntValue: Id {92156321-3e30-463a-83fa-c306bca1bc5c}
   Method FromULIntReference: Id {a686507f-51c4-410e-98ad-c2541ef602d2}
   Method FromULIntValue: Id {86c92bb6-733a-407c-aa95-3d976887e765}
   Method FromUSIntReference: Id {946118fe-852d-4783-9124-b28f9c5aa505}
   Method FromUSIntValue: Id {aeae6bc1-69d5-4f8e-bf8c-5456e7fca1c3}
   Method FromWordReference: Id {3a044499-0651-4e47-8802-27ec81f73705}
   Method FromWordValue: Id {cf646851-d26b-43e6-9a97-f0629adff38e}
   Method FromWStringReference: Id {ef6f17c2-c854-4bd1-98d9-b20dcef69d2f}
   Method FromWStringValue: Id {7495b560-9d45-42dd-b7ac-cea5caf03cd8}
   Property NamespaceName: Id {1b7a4363-1ae3-4082-9387-38baaafa2b6f}
   Get Get: Id {d9491450-ccd1-4cff-a47e-d13d4898b8f0} *)
